// TIA Portal V19 export
// export: Created 2000-01-01T00:00:00.0000000Z, ExportSetting None
FUNCTION "FC_Rung" : Void   // FC42, LAD
{ S7_Optimized_Access := 'TRUE' }
   VAR_INPUT
      Local : Int;
   END_VAR
BEGIN

REGION Network 1
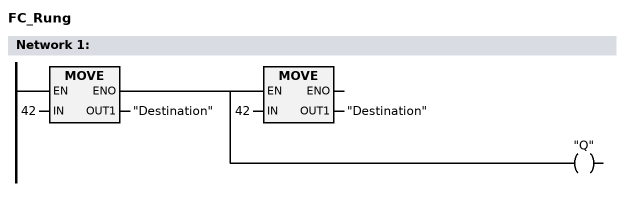
   RUNG wire#powerrail
      { S7_GenerateENO := "TRUE" } Move(in := 42, out1 => "Destination")
      wire#w1
      Move(in := 42, out1 => "Destination")
   END_RUNG
   RUNG wire#w1
      Coil( "Q" )
   END_RUNG
   // the same network as SCL:
   // ENO of a box is taken as its EN; it also drops when the box reports an error
   "Destination" := 42;
   "Destination" := 42;
   "Q" := TRUE;
END_REGION
END_FUNCTION
